Fanuc KAREL source: kt00749.KL

-- PROVISIONAL review KL for V1013-1; original PC SHA256 649474f50f6a48d1a0be96ba0012905c3a9c91fdd8b6f13e92a094736d3068fb
-- Incomplete behavior may be omitted. Consult companion uncertainty JSON. Do not deploy.
PROGRAM KT00749
%NOLOCKGROUP
VAR
  I1 : INTEGER
  I2 : INTEGER
  OUT : REAL
BEGIN
  -- UNRESOLVED_PC offsets 5-16; opcodes 2E,23
  -- UNRESOLVED_PC offsets 21-32; opcodes 2E,23
  -- UNRESOLVED_PC offsets 37-48; opcodes 2E,23
  -- UNRESOLVED_PC offsets 53-64; opcodes 2E,23
  -- UNRESOLVED_PC offsets 69-83; opcodes 21,50,64,23
  -- UNRESOLVED_PC offsets 88-92; opcodes 7F
END KT00749
